Fanuc KAREL source: compact_preamble.KL

PROGRAM KA00054
%NOLOCKGROUP
VAR
SRC : POSITION;DST : XYZWPR
BEGIN
DST=SRC
END KA00054
